// TwinCAT 3 PLC project PLC1
// ProgramVersion: 3.1.4026.27
// CompilerDefines: VISU_USEPROPERTYINFO
// libraries:
//   Tc2_Standard, * (Beckhoff Automation GmbH)
//   Tc2_System, * (Beckhoff Automation GmbH)
//   VisuSymbols, 4.5.0.0 (System)
// project tree:
//   / GlobalTextList.TcGTLO, PlcTask.TcTTO, Visualization Manager.TcVMO (not stored)
//   POUs/ MAIN.TcPOU
//   VISUs/ Visualization.TcVIS
// real-time tasks:
//   TASK PlcTask: cycle T#10ms, priority 20, ADS port 350

CONFIGURATION PLC1
    RESOURCE PLC ON TwinCAT3
        TASK PlcTask(INTERVAL := T#10ms, PRIORITY := 20);
        PROGRAM MAIN WITH PlcTask : MAIN;
    END_RESOURCE
END_CONFIGURATION

// ---- POUs/MAIN.TcPOU
PROGRAM MAIN
VAR
    //INPUTS
    iNumber   : INT;
    bSwitch1  : BOOL;
    bSwitch2  : BOOL;
    bSwitch3  : BOOL;
    bSwitch4  : BOOL;
    
    //OUTPUTS
    bLight1   : BOOL;
    bLight2   : BOOL;
    bLight3   : BOOL;
    bLight4   : BOOL;
END_VAR

bLight1 := bLight2 := bLight3 := bLight4 := FALSE;

IF (iNumber >= 0) AND (iNumber <= 8000) THEN
    bLight1 := TRUE;
ELSIF (iNumber > 8000) AND (iNumber <= 16000) THEN
    bLight2 := TRUE;
ELSIF (iNumber > 16000) AND (iNumber <= 24000) THEN
    bLight3 := TRUE;
ELSE
    bLight4 := TRUE;
END_IF

END_PROGRAM

// ---- GlobalTextList.TcGTLO
TEXTLIST GlobalTextList
  334 = '%i'
  838 = '%I.0'
  443 = 'iNumber'
  183 = 'Switch 1'
  127 = 'Switch 2'
  470 = 'Switch 3'
  294 = 'Switch 4'
END_TEXTLIST

// ---- VISUs/Visualization.TcVIS
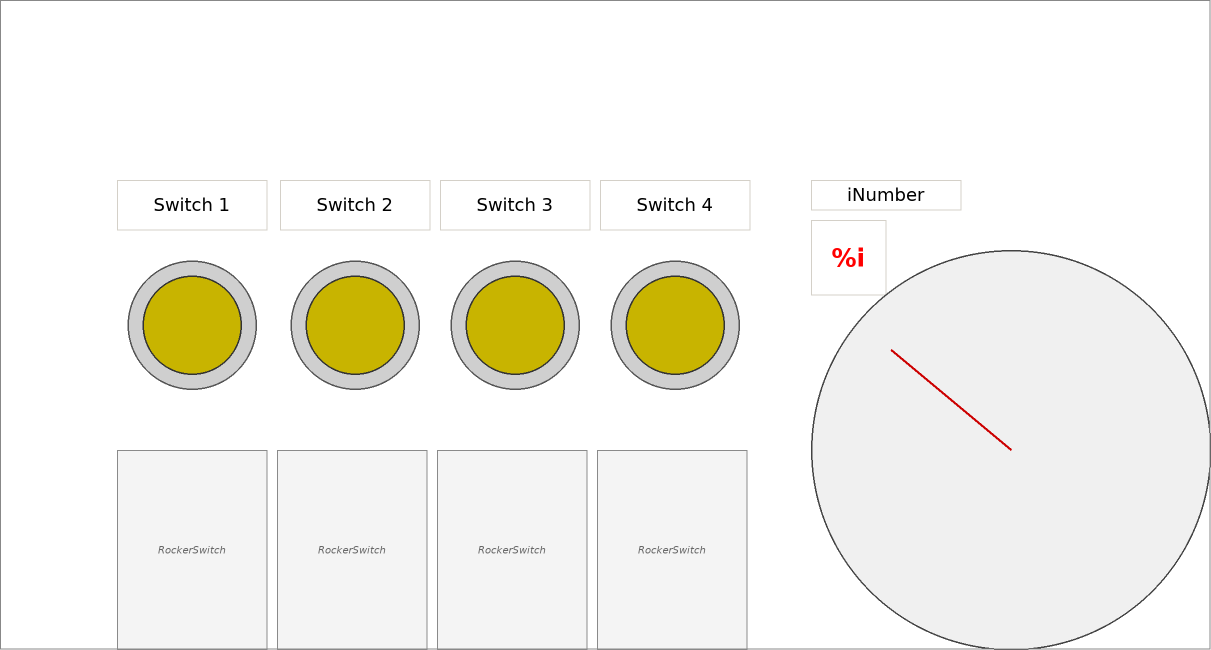
VISUALIZATION Visualization  // 1211x650
    RockerSwitch (117,450 150x200), variable: MAIN.bSwitch1, behaviour: TOGGLE, style: Switch-RockerSwitch-Gray
    RockerSwitch (277,450 150x200), variable: MAIN.bSwitch2, behaviour: TOGGLE, style: Switch-RockerSwitch-Gray
    RockerSwitch (437,450 150x200), variable: MAIN.bSwitch3, behaviour: TOGGLE, style: Switch-RockerSwitch-Gray
    RockerSwitch (597,450 150x200), variable: MAIN.bSwtich4, behaviour: TOGGLE, style: Switch-RockerSwitch-Gray
    Lamp1 (117,250 150x150), variable: MAIN.bLight1, style: Lamp-Lamp1-Yellow
    Lamp1 (440,250 150x150), variable: MAIN.bLight3, style: Lamp-Lamp1-Yellow
    Lamp1 (280,250 150x150), variable: MAIN.bLight2, style: Lamp-Lamp1-Yellow
    Lamp1 (600,250 150x150), variable: MAIN.bLight4, style: Lamp-Lamp1-Yellow
    Textfield (117,180 150x50), "Switch 1"
    Textfield (280,180 150x50), "Switch 2"
    Textfield (440,180 150x50), "Switch 3"
    Textfield (600,180 150x50), "Switch 4"
    Textfield (811,220 75x75), "%i", text variable: MAIN.iNumber
    Textfield (811,180 150x30), "iNumber"
    Meter360 (811,250 400x400), value: MAIN.iNumber, style: Meter-Meter360-Gray, scale format: %.1f, scale 0..32000
END_VISUALIZATION
